Fanuc KAREL source: compact_preamble.KL

PROGRAM KD00044
%NOLOCKGROUP
VAR
I:INTEGER;J:INTEGER;B:BOOLEAN;R:REAL;S : STRING[80]
-- UNRESOLVED DECLARATIONS (source type spelling not recovered)
-- G : TYPE_0x011E (type_u16=0x011E)
BEGIN
I=1
END KD00044
